// TIA Portal V21 export
FUNCTION_BLOCK "FB_AnaStatusIgnored"   // FB18, SCL
TITLE = Analyzer: status never evaluated
{ S7_Optimized_Access := 'TRUE' }
// Rule C26n: RET_VAL of RD_LOC_T is stored but never evaluated
// stored: MemoryReserve 100, SetENOAutomatically false
   VAR
      Now : DTL;   // Local time
   END_VAR
   VAR_TEMP
      RetVal : Int;   // Status of RD_LOC_T
   END_VAR
BEGIN

       #RetVal := RD_LOC_T(OUT => #Now);
END_FUNCTION_BLOCK
